(* IEC 61131-3 sources: STAR-PLC-Agent/results/raw/four_group_20261114/star_deepseek_v2/PUB008/generation/sim_00, 1 file *)

(* ---- test_program.st ---- *)
PROGRAM PLC_PRG
VAR
 BenchStep : UDINT := 0;
 BenchCalls : UDINT := 0;
 BenchDone : BOOL := FALSE;
 BenchUut0 : FB_Task;
 BenchUut1 : FB_Task;
 Binding_0_analogValues : ARRAY[1..4] OF INT;
 Binding_0_channels : ARRAY[1..4] OF ST_AnalogChannel;
 Binding_1_analogValues : ARRAY[1..5] OF INT;
 Binding_1_channels : ARRAY[1..5] OF ST_AnalogChannel;
 TraceIn_count : ARRAY[0..1] OF DINT;
 TraceOut_analogValues_1 : ARRAY[0..1] OF INT;
 TraceOut_analogValues_2 : ARRAY[0..1] OF INT;
 TraceOut_analogValues_3 : ARRAY[0..1] OF INT;
 TraceOut_analogValues_4 : ARRAY[0..1] OF INT;
 TraceOut_analogValues_5 : ARRAY[0..1] OF INT;
 TraceOut_channels_1_enable : ARRAY[0..1] OF BOOL;
 TraceOut_channels_1_hiLIM : ARRAY[0..1] OF REAL;
 TraceOut_channels_1_loLIM : ARRAY[0..1] OF REAL;
 TraceOut_channels_1_bipolar : ARRAY[0..1] OF BOOL;
 TraceOut_channels_1_measuringMode : ARRAY[0..1] OF INT;
 TraceOut_channels_1_retVal : ARRAY[0..1] OF WORD;
 TraceOut_channels_1_outputValue : ARRAY[0..1] OF REAL;
 TraceOut_channels_2_enable : ARRAY[0..1] OF BOOL;
 TraceOut_channels_2_hiLIM : ARRAY[0..1] OF REAL;
 TraceOut_channels_2_loLIM : ARRAY[0..1] OF REAL;
 TraceOut_channels_2_bipolar : ARRAY[0..1] OF BOOL;
 TraceOut_channels_2_measuringMode : ARRAY[0..1] OF INT;
 TraceOut_channels_2_retVal : ARRAY[0..1] OF WORD;
 TraceOut_channels_2_outputValue : ARRAY[0..1] OF REAL;
 TraceOut_channels_3_enable : ARRAY[0..1] OF BOOL;
 TraceOut_channels_3_hiLIM : ARRAY[0..1] OF REAL;
 TraceOut_channels_3_loLIM : ARRAY[0..1] OF REAL;
 TraceOut_channels_3_bipolar : ARRAY[0..1] OF BOOL;
 TraceOut_channels_3_measuringMode : ARRAY[0..1] OF INT;
 TraceOut_channels_3_retVal : ARRAY[0..1] OF WORD;
 TraceOut_channels_3_outputValue : ARRAY[0..1] OF REAL;
 TraceOut_channels_4_enable : ARRAY[0..1] OF BOOL;
 TraceOut_channels_4_hiLIM : ARRAY[0..1] OF REAL;
 TraceOut_channels_4_loLIM : ARRAY[0..1] OF REAL;
 TraceOut_channels_4_bipolar : ARRAY[0..1] OF BOOL;
 TraceOut_channels_4_measuringMode : ARRAY[0..1] OF INT;
 TraceOut_channels_4_retVal : ARRAY[0..1] OF WORD;
 TraceOut_channels_4_outputValue : ARRAY[0..1] OF REAL;
 TraceOut_channels_5_enable : ARRAY[0..1] OF BOOL;
 TraceOut_channels_5_hiLIM : ARRAY[0..1] OF REAL;
 TraceOut_channels_5_loLIM : ARRAY[0..1] OF REAL;
 TraceOut_channels_5_bipolar : ARRAY[0..1] OF BOOL;
 TraceOut_channels_5_measuringMode : ARRAY[0..1] OF INT;
 TraceOut_channels_5_retVal : ARRAY[0..1] OF WORD;
 TraceOut_channels_5_outputValue : ARRAY[0..1] OF REAL;
END_VAR

IF NOT BenchDone THEN
 CASE BenchStep OF
 0:
   Binding_0_analogValues[1] := INT#13824;
   Binding_0_analogValues[2] := INT#-13824;
   Binding_0_analogValues[3] := INT#1234;
   Binding_0_analogValues[4] := INT#5678;
   Binding_0_channels[1].enable := TRUE;
   Binding_0_channels[1].hiLIM := REAL#100.0;
   Binding_0_channels[1].loLIM := REAL#0.0;
   Binding_0_channels[1].bipolar := FALSE;
   Binding_0_channels[1].measuringMode := INT#0;
   Binding_0_channels[1].retVal := WORD#777;
   Binding_0_channels[1].outputValue := REAL#777.7;
   Binding_0_channels[2].enable := TRUE;
   Binding_0_channels[2].hiLIM := REAL#10.0;
   Binding_0_channels[2].loLIM := REAL#-10.0;
   Binding_0_channels[2].bipolar := TRUE;
   Binding_0_channels[2].measuringMode := INT#0;
   Binding_0_channels[2].retVal := WORD#777;
   Binding_0_channels[2].outputValue := REAL#777.7;
   Binding_0_channels[3].enable := TRUE;
   Binding_0_channels[3].hiLIM := REAL#100.0;
   Binding_0_channels[3].loLIM := REAL#0.0;
   Binding_0_channels[3].bipolar := FALSE;
   Binding_0_channels[3].measuringMode := INT#1;
   Binding_0_channels[3].retVal := WORD#777;
   Binding_0_channels[3].outputValue := REAL#777.7;
   Binding_0_channels[4].enable := TRUE;
   Binding_0_channels[4].hiLIM := REAL#100.0;
   Binding_0_channels[4].loLIM := REAL#0.0;
   Binding_0_channels[4].bipolar := FALSE;
   Binding_0_channels[4].measuringMode := INT#2;
   Binding_0_channels[4].retVal := WORD#777;
   Binding_0_channels[4].outputValue := REAL#777.7;
   BenchUut0.count := DINT#4;
   TraceIn_count[0] := BenchUut0.count;
   BenchUut0(analogValues := Binding_0_analogValues, channels := Binding_0_channels);
   TraceOut_analogValues_1[0] := Binding_0_analogValues[1];
   TraceOut_analogValues_2[0] := Binding_0_analogValues[2];
   TraceOut_analogValues_3[0] := Binding_0_analogValues[3];
   TraceOut_analogValues_4[0] := Binding_0_analogValues[4];
   TraceOut_channels_1_enable[0] := Binding_0_channels[1].enable;
   TraceOut_channels_1_hiLIM[0] := Binding_0_channels[1].hiLIM;
   TraceOut_channels_1_loLIM[0] := Binding_0_channels[1].loLIM;
   TraceOut_channels_1_bipolar[0] := Binding_0_channels[1].bipolar;
   TraceOut_channels_1_measuringMode[0] := Binding_0_channels[1].measuringMode;
   TraceOut_channels_1_retVal[0] := Binding_0_channels[1].retVal;
   TraceOut_channels_1_outputValue[0] := Binding_0_channels[1].outputValue;
   TraceOut_channels_2_enable[0] := Binding_0_channels[2].enable;
   TraceOut_channels_2_hiLIM[0] := Binding_0_channels[2].hiLIM;
   TraceOut_channels_2_loLIM[0] := Binding_0_channels[2].loLIM;
   TraceOut_channels_2_bipolar[0] := Binding_0_channels[2].bipolar;
   TraceOut_channels_2_measuringMode[0] := Binding_0_channels[2].measuringMode;
   TraceOut_channels_2_retVal[0] := Binding_0_channels[2].retVal;
   TraceOut_channels_2_outputValue[0] := Binding_0_channels[2].outputValue;
   TraceOut_channels_3_enable[0] := Binding_0_channels[3].enable;
   TraceOut_channels_3_hiLIM[0] := Binding_0_channels[3].hiLIM;
   TraceOut_channels_3_loLIM[0] := Binding_0_channels[3].loLIM;
   TraceOut_channels_3_bipolar[0] := Binding_0_channels[3].bipolar;
   TraceOut_channels_3_measuringMode[0] := Binding_0_channels[3].measuringMode;
   TraceOut_channels_3_retVal[0] := Binding_0_channels[3].retVal;
   TraceOut_channels_3_outputValue[0] := Binding_0_channels[3].outputValue;
   TraceOut_channels_4_enable[0] := Binding_0_channels[4].enable;
   TraceOut_channels_4_hiLIM[0] := Binding_0_channels[4].hiLIM;
   TraceOut_channels_4_loLIM[0] := Binding_0_channels[4].loLIM;
   TraceOut_channels_4_bipolar[0] := Binding_0_channels[4].bipolar;
   TraceOut_channels_4_measuringMode[0] := Binding_0_channels[4].measuringMode;
   TraceOut_channels_4_retVal[0] := Binding_0_channels[4].retVal;
   TraceOut_channels_4_outputValue[0] := Binding_0_channels[4].outputValue;
   BenchCalls := BenchCalls + 1;
 1:
   Binding_1_analogValues[1] := INT#5000;
   Binding_1_analogValues[2] := INT#100;
   Binding_1_analogValues[3] := INT#13824;
   Binding_1_analogValues[4] := INT#5678;
   Binding_1_analogValues[5] := INT#999;
   Binding_1_channels[1].enable := TRUE;
   Binding_1_channels[1].hiLIM := REAL#0.0;
   Binding_1_channels[1].loLIM := REAL#10.0;
   Binding_1_channels[1].bipolar := FALSE;
   Binding_1_channels[1].measuringMode := INT#3;
   Binding_1_channels[1].retVal := WORD#0;
   Binding_1_channels[1].outputValue := REAL#111.1;
   Binding_1_channels[2].enable := TRUE;
   Binding_1_channels[2].hiLIM := REAL#5.0;
   Binding_1_channels[2].loLIM := REAL#5.0;
   Binding_1_channels[2].bipolar := FALSE;
   Binding_1_channels[2].measuringMode := INT#1;
   Binding_1_channels[2].retVal := WORD#0;
   Binding_1_channels[2].outputValue := REAL#222.2;
   Binding_1_channels[3].enable := FALSE;
   Binding_1_channels[3].hiLIM := REAL#0.0;
   Binding_1_channels[3].loLIM := REAL#10.0;
   Binding_1_channels[3].bipolar := FALSE;
   Binding_1_channels[3].measuringMode := INT#9;
   Binding_1_channels[3].retVal := WORD#123;
   Binding_1_channels[3].outputValue := REAL#333.3;
   Binding_1_channels[4].enable := TRUE;
   Binding_1_channels[4].hiLIM := REAL#100.0;
   Binding_1_channels[4].loLIM := REAL#0.0;
   Binding_1_channels[4].bipolar := FALSE;
   Binding_1_channels[4].measuringMode := INT#2;
   Binding_1_channels[4].retVal := WORD#999;
   Binding_1_channels[4].outputValue := REAL#999.9;
   Binding_1_channels[5].enable := TRUE;
   Binding_1_channels[5].hiLIM := REAL#0.0;
   Binding_1_channels[5].loLIM := REAL#10.0;
   Binding_1_channels[5].bipolar := FALSE;
   Binding_1_channels[5].measuringMode := INT#9;
   Binding_1_channels[5].retVal := WORD#444;
   Binding_1_channels[5].outputValue := REAL#444.4;
   BenchUut1.count := DINT#4;
   TraceIn_count[1] := BenchUut1.count;
   BenchUut1(analogValues := Binding_1_analogValues, channels := Binding_1_channels);
   TraceOut_analogValues_1[1] := Binding_1_analogValues[1];
   TraceOut_analogValues_2[1] := Binding_1_analogValues[2];
   TraceOut_analogValues_3[1] := Binding_1_analogValues[3];
   TraceOut_analogValues_4[1] := Binding_1_analogValues[4];
   TraceOut_analogValues_5[1] := Binding_1_analogValues[5];
   TraceOut_channels_1_enable[1] := Binding_1_channels[1].enable;
   TraceOut_channels_1_hiLIM[1] := Binding_1_channels[1].hiLIM;
   TraceOut_channels_1_loLIM[1] := Binding_1_channels[1].loLIM;
   TraceOut_channels_1_bipolar[1] := Binding_1_channels[1].bipolar;
   TraceOut_channels_1_measuringMode[1] := Binding_1_channels[1].measuringMode;
   TraceOut_channels_1_retVal[1] := Binding_1_channels[1].retVal;
   TraceOut_channels_1_outputValue[1] := Binding_1_channels[1].outputValue;
   TraceOut_channels_2_enable[1] := Binding_1_channels[2].enable;
   TraceOut_channels_2_hiLIM[1] := Binding_1_channels[2].hiLIM;
   TraceOut_channels_2_loLIM[1] := Binding_1_channels[2].loLIM;
   TraceOut_channels_2_bipolar[1] := Binding_1_channels[2].bipolar;
   TraceOut_channels_2_measuringMode[1] := Binding_1_channels[2].measuringMode;
   TraceOut_channels_2_retVal[1] := Binding_1_channels[2].retVal;
   TraceOut_channels_2_outputValue[1] := Binding_1_channels[2].outputValue;
   TraceOut_channels_3_enable[1] := Binding_1_channels[3].enable;
   TraceOut_channels_3_hiLIM[1] := Binding_1_channels[3].hiLIM;
   TraceOut_channels_3_loLIM[1] := Binding_1_channels[3].loLIM;
   TraceOut_channels_3_bipolar[1] := Binding_1_channels[3].bipolar;
   TraceOut_channels_3_measuringMode[1] := Binding_1_channels[3].measuringMode;
   TraceOut_channels_3_retVal[1] := Binding_1_channels[3].retVal;
   TraceOut_channels_3_outputValue[1] := Binding_1_channels[3].outputValue;
   TraceOut_channels_4_enable[1] := Binding_1_channels[4].enable;
   TraceOut_channels_4_hiLIM[1] := Binding_1_channels[4].hiLIM;
   TraceOut_channels_4_loLIM[1] := Binding_1_channels[4].loLIM;
   TraceOut_channels_4_bipolar[1] := Binding_1_channels[4].bipolar;
   TraceOut_channels_4_measuringMode[1] := Binding_1_channels[4].measuringMode;
   TraceOut_channels_4_retVal[1] := Binding_1_channels[4].retVal;
   TraceOut_channels_4_outputValue[1] := Binding_1_channels[4].outputValue;
   TraceOut_channels_5_enable[1] := Binding_1_channels[5].enable;
   TraceOut_channels_5_hiLIM[1] := Binding_1_channels[5].hiLIM;
   TraceOut_channels_5_loLIM[1] := Binding_1_channels[5].loLIM;
   TraceOut_channels_5_bipolar[1] := Binding_1_channels[5].bipolar;
   TraceOut_channels_5_measuringMode[1] := Binding_1_channels[5].measuringMode;
   TraceOut_channels_5_retVal[1] := Binding_1_channels[5].retVal;
   TraceOut_channels_5_outputValue[1] := Binding_1_channels[5].outputValue;
   BenchCalls := BenchCalls + 1;
 END_CASE;
 BenchStep := BenchStep + 1;
 IF BenchStep >= 2 THEN BenchDone := TRUE; END_IF;
END_IF;
END_PROGRAM
